TYPE "ST_SignalTowerOut"
VERSION : 0.1
   STRUCT
      Red : Bool;
      Amber : Bool;
      Green : Bool;
      Blue : Bool;
      White : Bool;
      Horn : Bool;
      TestActive : Bool;
   END_STRUCT;

END_TYPE

